(* IEC 61131-3 sources: virtual-bottling-plant/plc/src/generated/gvl, 1 file *)

(* ---- GVL_Contract.st ---- *)
(* GENERATED by plc/scripts/gen_plc_io.py from contracts/modbus/sim-io.yaml + plc-io.yaml. Do not edit by hand. *)
(* Global process image. Only the generated IO_* / Bridge_* programs and PRG_Main use these. *)
  VAR_GLOBAL
    G_In : ST_SimInputs;
    G_Out : ST_SimOutputs;
    G_Status : ST_Status;
    G_Comms : ST_CommsStatus;
    G_Alarms : ST_AlarmSummary;
    G_Counters : ST_Counters;
    G_Cmd : ST_Commands;
    G_RecipeReq : ST_RecipeRequest;
    G_RecipeResp : ST_RecipeResponse;
  END_VAR
